// TIA Portal V17 export
// export: Created 2026-11-08T05:50:28.55177Z, ExportSetting WithDefaults, DisplayName Totally Integrated Automation Portal, DisplayVersion V17, DisplayName TIA Portal Openness, DisplayVersion V17, DisplayName TIA Portal Version Control Interface, DisplayVersion V17, DisplayName STEP 7 Professional, DisplayVersion V17, DisplayName STEP 7 Safety, DisplayVersion V17, DisplayName WinCC Professional, DisplayVersion V17
DATA_BLOCK "DB_HMI"   // DB1
{ S7_Optimized_Access := 'TRUE' }
VERSION : 0.1
// stored: AutoNumber true, DBAccessibleFromOPCUA true, IsOnlyStoredInLoadMemory false, IsRetainMemResEnabled false, IsWriteProtectedInAS false, MemoryReserve 100
   VAR
      Cmd_Marcha : Bool;   // Boton MARCHA de la HMI (momentaneo)
      Cmd_Paro : Bool;   // Boton PARO de la HMI (momentaneo)
      Cmd_Reset : Bool;   // Boton RESET de la HMI (momentaneo)
      Sel_Estilo : Int := 1;   // 1 Banderas, 2 Moore, 3 Mealy
      Estado : Int;   // Estado del estilo seleccionado: 0 Reposo, 10 Marcha, 90 Falla
      Motor_En_Marcha : Bool;   // Copia de KM1_Motor para la HMI
      Falla_Termico : Bool;   // Termico disparado
      Pantalla : Int;   // Pantalla activa en la HMI (1 Principal, 2 Diagnostico, 3 Estilos)
   END_VAR
BEGIN
END_DATA_BLOCK
